(* IEC 61131-3 sources: Versio-VersionControlSystem/fixtures/projects/RefrigeratorControl_FBS/RefrigeratorControl.fbsproj/Device.device.xml.v3^/Plc Logic.plclogic.xml.v3^/Application.application.xml.v3^, 3 files *)

(* ---- Glob_Var.gvl ---- *)
(* METADATA
{
	"v3Meta": {
		"objectGuid": "f8ccf7f9-314d-4201-b460-0f935fbcbf7d"
	}
}
*)
{attribute 'qualified_only'}
NAMESPACE Glob_Var
VAR_GLOBAL
//Inputs
	TempActual: REAL:=8.0;
	TempSet: REAL:=8.0;
	DoorOpen: BOOL;
	AlarmThreshold:TIME:=T#10S;
	DoorOpenThreshold:TIME:=T#10S;

//Outputs
	Compressor: BOOL;
	Signal: BOOL;
	Lamp: BOOL;
END_VAR
END_NAMESPACE

(* ---- PLC_PRG.prg.st ---- *)
(* METADATA
{
	"v3Meta": {
		"objectGuid": "e5cd9370-6160-4e13-a6ef-514133c47037"
	}
}
*)
PROGRAM PLC_PRG
VAR
	Alarm 		: FB_Alarm;
	Trigger 	: BOOL;
	OnTime		: TIME := T#2S;
	OffTime		: TIME := T#5S;
	Latch		: BOOL := FALSE;
END_VAR

Alarm.P_Settings.Latch := Latch;
Alarm.P_Settings.OnDelayTime := OnTime;
Alarm.P_Settings.OffDelayTime := OffTime;
Alarm.Condition := Trigger;
Alarm();
END_PROGRAM

(* ---- Simulation.prg.st ---- *)
(* METADATA
{
	"v3Meta": {
		"objectGuid": "980a4bef-b0b7-4f16-816b-1f41192a0ee0"
	}
}
*)
PROGRAM Simulation
VAR
	T1: TON;					//The temperature is decreased on a time delay, when the comepressor has been activated
	P_Cooling: TIME:=T#500MS;
	xReduceTemp: BOOL;			//Signal for dereasing the temperature
	T2: TON;					//The temperature is increased on a time delay, when the compressor has been activated
	P_Environment: TIME:=T#2S;			//Delay time when the door is closed
	P_EnvironmentDoorOpen: TIME:=T#1S;	//Delay time when the door is open
	xRaiseTemp: BOOL;					//Signal for increasing the temperature
	tTemp: TIME;						//Delay time
	TestTag : BOOL;
	TestTAg2: BOOL;
END_VAR

// After the compressor has been activated due to TempActual being too high, the temperature decreases.
// The temperature is decremented by 0.1°C per cycle after a delay of P_Cooling
IF Glob_Var.Compressor THEN
	T1(IN:= Glob_Var.Compressor, PT:= P_Cooling, Q=>xReduceTemp);
	IF xReduceTemp THEN
		Glob_Var.TempActual := Glob_Var.TempActual-0.1;
		T1(IN:=FALSE);
	END_IF
END_IF

//If the door is open, the warming occurs faster; SEL selects P_EnvironmentDoorOpen
tTemp:=SEL(Glob_Var.DoorOpen, P_Environment, P_EnvironmentDoorOpen);

//If the compressor is not in operation, then the cooling chamber becomes warmer.
//The  temperature is incremented by 0.1°C per cycle after a delay of tTemp
T2(IN:= TRUE, PT:= tTemp, Q=>xRaiseTemp);
IF xRaiseTemp THEN
	Glob_Var.TempActual := Glob_Var.TempActual + 0.1;
	T2(IN:=FALSE);
END_IF
END_PROGRAM
